TYPE ST_PolarIIChamber_ChamberServiceCtrl :
STRUCT
	SetMode : ST_ServiceCtrl;
	Initial : ST_ServiceCtrl;
	SingleProcess : ST_ServiceCtrl;
	EMGS : ST_ServiceCtrl;
	SetConfig : ST_ServiceCtrl;
	ArmAlignTest : ST_ServiceCtrl;
	ArmTest : ST_ServiceCtrl;
	FlowCalibration : ST_ServiceCtrl;
	CupChamberClean : ST_ServiceCtrl;
	DoNozzleClean : ST_ServiceCtrl;
	DoNozzlePreflush : ST_ServiceCtrl;
END_STRUCT
END_TYPE

(* stored: Version 1.1.0.1, ProductVersion 3.1.4026.18
   DUT ST_PolarIIChamber_ChamberServiceCtrl: Id {14000000-0000-0000-0000-000000000019} *)
